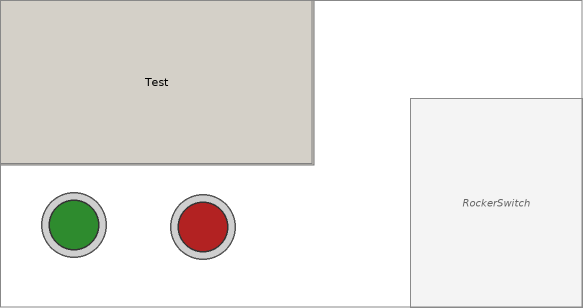
VISUALIZATION vis_Desolve  // 583x308
    Button (0,0 314x165), "Test"
    RockerSwitch (410,98 173x210), variable: gIO.q_EL[1].q_ch2, behaviour: TOGGLE, style: Switch-RockerSwitch-Red
    Lamp1 (36,186 76x78), style: Lamp-Lamp1-Green
    Lamp1 (165,188 76x78), style: Lamp-Lamp1-Red
END_VISUALIZATION

(* stored: Version 1.1.0.1, ProductVersion 3.1.4024.12
   Visu vis_Desolve: Id {a1332be3-adb7-4da6-a28e-5664dafe4728} *)
